Fanuc KAREL source: kt00893.compact.KL

PROGRAM KT00893
%STACKSIZE=65535
%PRIORITY=65535
%NOLOCKGROUP
VAR
P1 : POSITION
P2 : POSITION
OUT : BOOLEAN
BEGIN
OUT=IN_RANGE(P1)
END KT00893
